(* IEC 61131-3 sources: codesys-framework/txt/application/WeVe Utils (library)/TimeStamp/FB_TimeStampService/Utilities, 4 files *)

(* ---- GetLocalTime.method.st ---- *)
METHOD PRIVATE GetLocalTime : E_TaskStatus;
VAR_INPUT
END_VAR

// --- BEGIN IMPLEMENTATION ---

GetLocalTime := ReadParameter(
	wIndex			:= 16#245C,
	bySubIndex		:= 2,
	udiTimeOut		:= 1000,
	pDataBuffer		:= ADR(_uliParRead),
	udiBufferSize	:= 8
);

IF GetLocalTime = E_TaskStatus.Successful THEN
	_dtRead	:= ULINT_TO_DT(_uliParRead/1000000000+946684800);  //Compensation for 1/1/1970 vs 1/1/2000
	_sTimeStamp_Local_AsString := CONCAT (STR1 := RIGHT (STR := DT_TO_STRING (_dtRead), SIZE := 19), STR2 := '.000');
END_IF

(* ---- GetSystemTime_UTC.method.st ---- *)
METHOD PRIVATE GetSystemTime_UTC : BOOL
VAR_INPUT
END_VAR

// --- BEGIN IMPLEMENTATION ---

// Get SystemTime (UTC)
_fbGetSystemTime_UTC (xExecute := _xGetSystemTime, dtDateAndTime => _dtSystemTime_UTC);
_xGetSystemTime := TRUE;

IF _fbGetSystemTime_UTC.xDone THEN
	_xGetSystemTime := FALSE;
END_IF

// String of the UTC-DateTime
IF _fbGetSystemTime_UTC.xDone THEN
	_sTimeStamp_UTC_AsString := CONCAT(STR1 := RIGHT (STR := DT_TO_STRING (_dtSystemTime_UTC), SIZE := 19), STR2 := '.000');
	_xTimeStampStringCreated := TRUE;
END_IF

(* ---- ReadParameter.method.st ---- *)
METHOD PRIVATE ReadParameter : E_TaskStatus
VAR_INPUT
	wIndex				: WORD;
	bySubIndex			: BYTE;
	udiTimeOut			: UDINT;
	pDataBuffer			: POINTER TO BYTE;
	udiBufferSize		: UDINT;
END_VAR

// --- BEGIN IMPLEMENTATION ---

ReadParameter := E_TaskStatus.Busy;

_fbL_IPAP_ParameterRead(
	xExecute		:=_xReadparameter ,
	xAbort			:= ,
	wIndex			:= wIndex,
	bySubIndex		:= bySubIndex,
	udiTimeOut		:= udiTimeOut,
	pDataBuffer		:= pDataBuffer,
	udiBufferSize	:= udiBufferSize,
	xDone			=> ,
	xBusy			=> ,
	xAborted		=> ,
	xError			=> ,
	eErrorId		=> ,
	udiDataRead		=> ,
	eDataType		=>
);

// Get LocalTime
CASE _wReadParameterState OF

	0 :
		_xReadparameter := TRUE;
		_wReadParameterState := _wReadParameterState + 10;

	10:
		IF _fbL_IPAP_ParameterRead.xDone THEN
			_wReadParameterState := _wReadParameterState + 10;
		END_IF

		IF _fbL_IPAP_ParameterRead.xError THEN
			_xReadparameter := FALSE;
			_wReadParameterState := 100;
		END_IF

	20:
		_xReadparameter := FALSE;
		_wReadParameterState := _wReadParameterState + 10;

	30:
		//Extra state to disable the FB
		_wReadParameterState := 0;
		ReadParameter := E_TaskStatus.Successful;

	100:
		_wReadParameterState := 0;
		ReadParameter := E_TaskStatus.Failed;

END_CASE

(* ---- WriteParameter.method.st ---- *)
METHOD PRIVATE WriteParameter : E_TaskStatus
VAR_INPUT
	wIndex				: WORD;
	bySubIndex			: BYTE;
	udiTimeOut			: UDINT;
	pDataBuffer			: POINTER TO BYTE;
	udiDataSize			: UDINT;
END_VAR

// --- BEGIN IMPLEMENTATION ---

WriteParameter := E_TaskStatus.Busy;

_fbL_IPAP_ParameterWrite(
	xExecute	:=_xWriteParameter,
	xAbort		:= ,
	wIndex		:= wIndex,
	bySubIndex	:= bySubIndex,
	udiTimeOut	:= udiTimeOut,
	pDataBuffer	:= pDataBuffer,
	udiDataSize	:= udiDataSize,
	xDone		=> ,
	xBusy		=> ,
	xAborted	=> ,
	xError		=> ,
	eErrorId	=>
);

CASE _wWriteParameterState OF

	0 :
		_xWriteParameter   := TRUE;
		_wWriteParameterState := _wWriteParameterState + 10;

	10:
		IF _fbL_IPAP_ParameterWrite.xDone THEN
			_xWriteParameter := FALSE;
			_wWriteParameterState := _wWriteParameterState + 10;
		END_IF

		IF _fbL_IPAP_ParameterWrite.xError THEN
			_xWriteParameter := FALSE;
			_wWriteParameterState := 100;
		END_IF

	20:
		//Extra state to disable the FB
		_wWriteParameterState := 0;
		WriteParameter := E_TaskStatus.Successful;

	100:
		_wWriteParameterState := 0;
		WriteParameter := E_TaskStatus.Failed;

END_CASE
